(* PLC project g_compressor_cycle, Anonymous Benchmark Suite 1.0 *)
(* stored: creationDateTime 2026-08-28T00:00:00 *)

PROGRAM g_compressor_cycle
  VAR_INPUT
    PressLow : BOOL;
    PressHigh : BOOL;
    MinOffDone : BOOL;
  END_VAR
  VAR_OUTPUT
    Load : BOOL;
  END_VAR

(* LD diagram, written out as Structured Text *)
Load := (Load OR PressLow AND MinOffDone) AND NOT PressHigh;
END_PROGRAM

CONFIGURATION Config0
  RESOURCE Res0 ON PLC
    TASK tcyclic(INTERVAL := T#10ms, PRIORITY := 0);
    PROGRAM inst0 WITH tcyclic : g_compressor_cycle;
  END_RESOURCE
END_CONFIGURATION
